{region 'Documentation'}
(*!
<summary>Checks whether the ULINT value is outside the inclusive range.</summary>
<description>

Minimum &gt; Maximum reports Error during active evaluation; equal bounds are
valid.

</description>
*)
{endregion}
FUNCTION_BLOCK AssertNotInRange_ULInt EXTENDS AssertionBase
VAR_INPUT
    IN : ULINT; //! Actual value checked or observed by this Assertion.
    Minimum : ULINT; //! Inclusive lower bound of the comparison; for a range, must not exceed Maximum.
    Maximum : ULINT; //! Inclusive upper bound of the comparison; for a range, must not be below Minimum.
END_VAR

SUPER^();

{region 'Documentation'}
(*!
<summary>Check whether the ULINT value is outside the inclusive range.</summary>
*)
{endregion}
METHOD PROTECTED Assert
VAR
    Message : STRING(GVL_Constants.MessageLength);
    MinimumText : STRING(GVL_Constants.AssertionValueLength);
    MaximumText : STRING(GVL_Constants.AssertionValueLength);
    ActualText : STRING(GVL_Constants.AssertionValueLength);
END_VAR
IF NOT EvaluationActive THEN
    RETURN;
END_IF;

IF Result = E_Result.Error THEN
    RETURN;
END_IF;

IF Minimum > Maximum THEN
    MinimumText := ULINT_TO_STRING(Minimum);
    MaximumText := ULINT_TO_STRING(Maximum);
    Message := CONCAT('Assertion error: minimum exceeds maximum. Minimum = ',
        MinimumText);
    Message := CONCAT(Message, ', Maximum = ');
    Message := CONCAT(Message, MaximumText);
    Message := CONCAT(Message, '.');
    Error(Message := Message);
    RETURN;
END_IF;

IF Result = E_Result.Failed THEN
    RETURN;
END_IF;

IF (IN >= Minimum) AND (IN <= Maximum) THEN
    MinimumText := ULINT_TO_STRING(Minimum);
    MaximumText := ULINT_TO_STRING(Maximum);
    ActualText := ULINT_TO_STRING(IN);
    Message := CONCAT('Assertion failed: value is inside forbidden range. Minimum = ',
        MinimumText);
    Message := CONCAT(Message, ', Maximum = ');
    Message := CONCAT(Message, MaximumText);
    Message := CONCAT(Message, ', Actual = ');
    Message := CONCAT(Message, ActualText);
    Message := CONCAT(Message, '.');
    Fail(Message := Message);
    RETURN;
END_IF;

Pass();
END_METHOD

END_FUNCTION_BLOCK

(* stored: Version 1.1.0.1
   POU AssertNotInRange_ULInt: Id {19f26d84-8e92-484e-8a24-bea2013abe8c}, SpecialFunc None
   Folder Internal: Id {39b6b918-42a4-45a7-9bfc-8559a34a2e50}
   Method Assert: Id {c6d7f817-03c8-4c19-b61b-cf0608840df8} *)
